(* IEC 61131-3 sources: plcassist-cli/packages/volt-lsp-iec/test-corpus/bakon-nano/Device/Plc Logic/Application/Library Manager/L_TP2P_TechModulesProcessFunctions, 25 files *)

(* ---- GETBOOLEANPROPERTY.fun ---- *)
FUNCTION GETBOOLEANPROPERTY : BOOL
VAR_INPUT
	STKEY : WSTRING;
END_VAR
END_FUNCTION

(* ---- GETCOMPANY.fun ---- *)
FUNCTION GETCOMPANY : WSTRING
END_FUNCTION

(* ---- GETNUMBERPROPERTY.fun ---- *)
FUNCTION GETNUMBERPROPERTY : DINT
VAR_INPUT
	STKEY : WSTRING;
END_VAR
END_FUNCTION

(* ---- GETTEXTPROPERTY.fun ---- *)
FUNCTION GETTEXTPROPERTY : WSTRING
VAR_INPUT
	STKEY : WSTRING;
END_VAR
END_FUNCTION

(* ---- GETTEXTPROPERTY2.fun ---- *)
FUNCTION GETTEXTPROPERTY2 : POINTER TO WSTRING
VAR_INPUT
	STKEY : WSTRING;
END_VAR
END_FUNCTION

(* ---- GETTITLE.fun ---- *)
FUNCTION GETTITLE : WSTRING
END_FUNCTION

(* ---- GETVERSION.fun ---- *)
FUNCTION GETVERSION : VERSION
END_FUNCTION

(* ---- GETVERSIONPROPERTY.fun ---- *)
FUNCTION GETVERSIONPROPERTY : VERSION
VAR_INPUT
	STKEY : WSTRING;
END_VAR
END_FUNCTION

(* ---- L_TP2P_TC_CELSIUSTOFAHRENHEIT_ABS.fun ---- *)
FUNCTION L_TP2P_TC_CELSIUSTOFAHRENHEIT_ABS : LREAL
VAR_INPUT
	LRINVAL : LREAL;
END_VAR
END_FUNCTION

(* ---- L_TP2P_TC_CELSIUSTOFAHRENHEIT_REL.fun ---- *)
FUNCTION L_TP2P_TC_CELSIUSTOFAHRENHEIT_REL : LREAL
VAR_INPUT
	LRINVAL : LREAL;
END_VAR
END_FUNCTION

(* ---- _TM_COMMONBASE.fb ---- *)
FUNCTION_BLOCK _TM_COMMONBASE EXTENDS L_TB2P_TM_Base
VAR
	XTMSTOP : BOOL;
	LWTCHECKSUM : LWORD;
	ERRORHANDLER : L_IE1P_ErrorHandler;
	PINPUTBASE : POINTER TO L_TP2P_TemperatureControlBaseIn;
	POUTPUTBASE : POINTER TO L_TP2P_TemperatureControlBaseOut;
END_VAR
END_FUNCTION_BLOCK

METHOD CALL_ALLOCPOINTADR
END_METHOD

METHOD CALL_CHECKREQUESTS
END_METHOD

METHOD CALL_CTRLREQACTIVE : BOOL
END_METHOD

METHOD CALL_OUTPUT
END_METHOD

METHOD CALL_REQUESTS_EXT
END_METHOD

METHOD CALL_RESETCOMMANDS
END_METHOD

METHOD CALL_RESETOUTPUT
END_METHOD

METHOD CALL_RESETSETERROR
END_METHOD

METHOD CALL_SETERROR
END_METHOD

METHOD CALL_STOP
END_METHOD

METHOD CALL_TMFUNCTIONALITY
END_METHOD

METHOD CALL_S000_CYCLIC
END_METHOD

METHOD CALL_S001_INIT
END_METHOD

METHOD CALL_S002_READY
END_METHOD

METHOD CALL_S996_STOP
END_METHOD

METHOD CALL_STATEMACHINE
END_METHOD

METHOD CALL_T000_ALLSTATES
END_METHOD

METHOD CALL_T002_READY
END_METHOD

METHOD CALL_S000_CYCLIC_OUT
END_METHOD

METHOD CALL_S999_ERROR_OUT
END_METHOD

METHOD CALL_STATEMACHINE_OUT
END_METHOD

METHOD CALL_T000_ALLSTATES_OUT
END_METHOD

(* ---- _TM_TEMPERATURECONTROLBASE.fb ---- *)
FUNCTION_BLOCK _TM_TEMPERATURECONTROLBASE EXTENDS _TM_CommonBase
VAR_OUTPUT
	PPAR : POINTER TO _scPar_TM_TemperatureControlBase;
	PSF : POINTER TO _scSF_TM_TemperatureControlBase;
	PAP : POINTER TO _scAP_TM_TemperatureControlBase;
END_VAR
VAR_IN_OUT
	SCPERSISTENTDATA : L_TP2P_scPD_TemperatureControlBase;
END_VAR
VAR
	TM_TEMPERATURECONTROLCONFIG : L_TB2P_ModuleHandlerConfig;
	PINPUT : POINTER TO L_TP2P_TemperatureControlBaseIn;
	POUTPUT : POINTER TO L_TP2P_TemperatureControlBaseOut;
	_PSCPARVISU : POINTER TO _scPar_TM_TemperatureControlBase;
	SCPD_ACT : REFERENCE TO L_TP2P_scPD_TemperatureControlBase;
	LRTASKCYCLE : LREAL := 0.01;
	XNOREGULATIONPARAM : BOOL := FALSE;
	FB_TASKINFO : L_TP2P_TC_GetTaskInfo;
	FB_TEMPSETFILTER : L_TP2P_TC_TempSetFilter;
	FB_TEMPACTPROCESSING : L_TP2P_TC_TempActProcessing;
	FB_MONITORING : L_TP2P_TC_Monitoring;
	FB_PIDCONTROLLER : L_TP2P_TC_PIDController;
	FB_PARAMETERSWITCHING : L_TP2P_TC_ParameterSwitching;
	FB_PWM : L_TP2P_TC_PWM;
	FB_DIFFCTRL : L_TP2P_TC_DiffCtrl;
	FB_PARAMETERIDENTIFICATION : L_TP2P_TC_ParameterIdentification;
	SCIDENTDIAG : _sc_TM_TC_IdentDiagInfo;
END_VAR
END_FUNCTION_BLOCK

METHOD CALL_ALLOCPOINTADR
END_METHOD

METHOD CALL_CTRLREQACTIVE : BOOL
END_METHOD

METHOD CALL_ERRORHANDLER
END_METHOD

METHOD CALL_INITDONE
END_METHOD

METHOD CALL_INITROUTINE
END_METHOD

METHOD CALL_INTERNALCTRL
END_METHOD

METHOD CALL_OUTPUT
END_METHOD

METHOD CALL_OUTPUT_SF
END_METHOD

METHOD CALL_REQUESTS_EXT
END_METHOD

METHOD CALL_RESETCOMMANDS
END_METHOD

METHOD CALL_RESETOUTPUT
END_METHOD

METHOD CALL_FBMETHODS
END_METHOD

METHOD CALL_FB_DIFFCTRL
END_METHOD

METHOD CALL_FB_DIFFCTRLINPUTS
END_METHOD

METHOD CALL_FB_MONITORING
END_METHOD

METHOD CALL_FB_MONITORINGINPUTS
END_METHOD

METHOD CALL_FB_PIDCONTROLLER
END_METHOD

METHOD CALL_FB_PIDCONTROLLERINPUTS
END_METHOD

METHOD CALL_FB_PWM
END_METHOD

METHOD CALL_FB_PWMINPUTS
END_METHOD

METHOD CALL_FB_PARAMETERIDENTIFICATION
END_METHOD

METHOD CALL_FB_PARAMETERIDENTIFICATIONINPUTS
END_METHOD

METHOD CALL_FB_PARAMETERSWITCHING
END_METHOD

METHOD CALL_FB_PARAMETERSWITCHINGINPUTS
END_METHOD

METHOD CALL_FB_TEMPACTPROCESSING
END_METHOD

METHOD CALL_FB_TEMPACTPROCESSINGINPUTS
END_METHOD

METHOD CALL_FB_TEMPSETFILTER
END_METHOD

METHOD CALL_FB_TEMPSETFILTERINPUTS
END_METHOD

METHOD CALL_S000_CYCLIC
END_METHOD

METHOD CALL_S002_READY
END_METHOD

METHOD CALL_S210_CONTROL
END_METHOD

METHOD CALL_S211_REGULATION
END_METHOD

METHOD CALL_S212_IDENTIFICATION
END_METHOD

METHOD CALL_S996_STOP
END_METHOD

METHOD CALL_STATEMACHINE
END_METHOD

METHOD CALL_T002_READY
END_METHOD

(* ---- GLOBALTEXTLIST.fb ---- *)
FUNCTION_BLOCK GLOBALTEXTLIST
VAR
	M_TEXTLISTFILE : STRING(255);
	_STNAMESPACE : STRING;
END_VAR
END_FUNCTION_BLOCK

(* ---- L_TP2P_TC_DIFFCTRL.fb ---- *)
FUNCTION_BLOCK L_TP2P_TC_DIFFCTRL
VAR_INPUT
	LRTASKCYCLE : LREAL := 0.001;
	XENABLE : BOOL;
	LRCONTROLVALUE : LREAL;
END_VAR
VAR_OUTPUT
	XDIFFPOSITIVEOUT : BOOL;
	XDIFFNEGATIVEOUT : BOOL;
END_VAR
VAR_IN_OUT
	SCPAR : _scPar_TM_TemperatureControlBase;
END_VAR
VAR
	LRSIMUCONTROL_PCT : LREAL := 0.0;
	LRCTRLDIFF_PCT : LREAL;
	LRTIME_100PCT : LREAL := 0;
	LRTIME_0PCT : LREAL := 0;
	LRMINIMALONTIME_S : LREAL := 1;
	LRMINIMALOFFTIME_S : LREAL := 1;
	LRACTUALONTIME_POSITIVE_S : LREAL := 0;
	LRACTUALOFFTIME_POSITIVE_S : LREAL := 0;
	LRACTUALONTIME_NEGATIVE_S : LREAL := 0;
	LRACTUALOFFTIME_NEGATIVE_S : LREAL := 0;
	XPOSOUTLAST : BOOL := FALSE;
	XNEGOUTLAST : BOOL := FALSE;
END_VAR
END_FUNCTION_BLOCK

(* ---- L_TP2P_TC_GETTASKINFO.fb ---- *)
FUNCTION_BLOCK L_TP2P_TC_GETTASKINFO
VAR_OUTPUT
	DWCYCLETIME : DWORD;
	LRCYCLETIME : LREAL;
END_VAR
VAR
	XFIRSTCYCLE : BOOL := TRUE;
	HANDLE : RTS_IEC_HANDLE;
	INTERVAL : UDINT;
END_VAR
END_FUNCTION_BLOCK

(* ---- L_TP2P_TC_MONITORING.fb ---- *)
FUNCTION_BLOCK L_TP2P_TC_MONITORING
VAR_INPUT
	LRTASKCYCLE : LREAL := 0.001;
	XENABLE : BOOL := FALSE;
	LRSETTEMP : LREAL := 0;
	LRACTTEMP : LREAL := 0;
	LRACTTEMPUNFILTERED : LREAL := 0;
END_VAR
VAR_OUTPUT
	XTEMPMAXCRITICALABSOLUTE : BOOL;
	XSETTEMPREACHED : BOOL;
	XTEMPMIN : BOOL;
	XTEMPMAX : BOOL;
	XSENSORMONITORINGVALUEMIN : BOOL;
	XSENSORMONITORINGVALUEMAX : BOOL;
	XSENSORMONITORINGCHANGEMAX : BOOL;
END_VAR
VAR_IN_OUT
	SCPAR : _scPar_TM_TemperatureControlBase;
END_VAR
VAR
	LRSETACTDIFF : LREAL;
	LRACTTEMPLASTCYCLE : LREAL;
	RTENABLE : R_TRIG;
END_VAR
END_FUNCTION_BLOCK

(* ---- L_TP2P_TC_PARAMETERIDENTIFICATION.fb ---- *)
FUNCTION_BLOCK L_TP2P_TC_PARAMETERIDENTIFICATION
VAR_INPUT
	XENABLE : BOOL := FALSE;
	LRTASKCYCLE : LREAL := 0.001;
	LRTEMPACT : LREAL;
END_VAR
VAR_OUTPUT
	XDONE : BOOL;
	XBUSY : BOOL;
	WERRORID : WORD;
	WSTEP : WORD;
	WPHASE : WORD;
	LRCONTROLVALUEOUT : LREAL;
	LRTAUDEAD : LREAL;
	LRKI : LREAL;
	LRIDENTS1ELAPSEDTIME : LREAL;
	LRIDENTS1TEMPACTGRADIENT : LREAL;
	LRIDENTS2TEMPSTART : LREAL;
	LRIDENTS2ELAPSEDTIME : LREAL;
	LRIDENTS2TEMPACTGRADIENT : LREAL;
	LRIDENTS3TAUDEADACT : LREAL;
	LRIDENTS3TAUDEADMAX : LREAL;
END_VAR
VAR_IN_OUT
	SCPAR : _scPar_TM_TemperatureControlBase;
	SCPD : L_TP2P_scPD_TemperatureControlBase;
	SCIDENTDIAG : _sc_TM_TC_IdentDiagInfo;
END_VAR
VAR
	DWREGDATASIZE : DWORD := 20;
	FB_TEMPACTT1 : L_TP2P_TC_PT1Process;
	LRTEMPACTVALUE : LREAL;
	LRTEMPACTGRADIENT : LREAL;
	LRTEMPACTLASTCYCLE : LREAL;
	LRTIMESTART_S1 : LREAL;
	LRTEMPSTART_S2 : LREAL;
	LRTIMESTART_S2 : LREAL;
	LRTEMPSTART_S3 : LREAL;
	LRTIMESTART_S3 : LREAL;
	LRCONTROLVALUESTART_S3 : LREAL;
	LRCONTROLVALUESTEP_S3 : LREAL;
	DICYCLECOUNT_S3 : DINT;
	UDIREG_N : UDINT;
	LRREG_SUMX : LREAL;
	LRREG_SUMY : LREAL;
	LRREG_SUMXX : LREAL;
	LRREG_SUMXY : LREAL;
	LRREG_XM : LREAL;
	LRREG_YM : LREAL;
	LRREG_A : LREAL;
	LRREG_B : LREAL;
	LRZAEHLER_B : LREAL;
	LRNENNER_B : LREAL;
	LRTAUDEADMAX : LREAL;
	LRTAUDEADACT : LREAL;
	LRBMAX : LREAL;
	LRPAR_STEP1TEMPCHANGEMAX : LREAL;
	LRPAR_STEP2CONTROLSTEPPCT : LREAL;
	LRPAR_STEP2TEMPCHANGEMAX : LREAL;
	LRPAR_STEP2TEMPDIFFMIN : LREAL;
	LRPAR_STEP2WAITTIMEMIN : LREAL;
	LRPAR_STEP2CONTROLVALUEMAXPCT : LREAL;
	LRPAR_STEP3CONTROLSTEPPCT : LREAL;
	LRPAR_STEP3TEMPDIFFMIN : LREAL;
	LRPAR_STEP3REGRESSIONTIME : LREAL;
	ALRXVAL : ARRAY [1..dwRegDataSize] OF LREAL;
	ALRYVAL : ARRAY [1..dwRegDataSize] OF LREAL;
	DWCNT : DWORD;
	XPERFORMCALCREGRESSION : BOOL := FALSE;
	LRR01 : LREAL;
	LRSAMPLETIME : LREAL := 0.1;
	LRBUFFERLENGTH : LREAL := 0;
END_VAR
END_FUNCTION_BLOCK

METHOD ADDREGPOINT
VAR_INPUT
	LRX : LREAL;
	LRY : LREAL;
END_VAR
END_METHOD

METHOD CALCREGRESSION
END_METHOD

METHOD PREPAREREGBUFFER
END_METHOD

METHOD RESET : BOOL
END_METHOD

(* ---- L_TP2P_TC_PARAMETERIDENTIFICATION_T30.fb ---- *)
FUNCTION_BLOCK L_TP2P_TC_PARAMETERIDENTIFICATION_T30
VAR_INPUT
	XENABLE : BOOL := FALSE;
	LRTASKCYCLE : LREAL := 0.001;
	LRTEMPACT : LREAL;
END_VAR
VAR_OUTPUT
	XDONE : BOOL;
	XBUSY : BOOL;
	WERRORID : WORD;
	WSTEP : WORD;
	WPHASE : WORD;
	LRCONTROLVALUEOUT : LREAL;
	LRTAUDEAD : LREAL;
	LRKI : LREAL;
END_VAR
VAR_IN_OUT
	SCPAR : _scPar_TM_TemperatureControlBase;
	SCPD : L_TP2P_scPD_TemperatureControlBase;
END_VAR
VAR
	DWREGDATASIZE : DWORD := 30;
	FB_TEMPACTT1 : L_TP2P_TC_PT1Process;
	LRTEMPACTVALUE : LREAL;
	LRTEMPACTGRADIENT : LREAL;
	LRTEMPACTLASTCYCLE : LREAL;
	LRTIMESTART_S1 : LREAL;
	LRTEMPSTART_S2 : LREAL;
	LRTIMESTART_S2 : LREAL;
	LRTEMPSTART_S3 : LREAL;
	LRTIMESTART_S3 : LREAL;
	LRCONTROLVALUESTART_S3 : LREAL;
	LRCONTROLVALUESTEP_S3 : LREAL;
	DICYCLECOUNT_S3 : DINT;
	UDIREG_N : UDINT;
	LRREG_SUMX : LREAL;
	LRREG_SUMY : LREAL;
	LRREG_SUMXX : LREAL;
	LRREG_SUMXY : LREAL;
	LRREG_XM : LREAL;
	LRREG_YM : LREAL;
	LRREG_A : LREAL;
	LRREG_B : LREAL;
	LRZAEHLER_B : LREAL;
	LRNENNER_B : LREAL;
	LRTAUDEADMAX : LREAL;
	LRTAUDEADACT : LREAL;
	LRBMAX : LREAL;
	LRPAR_STEP1TEMPCHANGEMAX : LREAL;
	LRPAR_STEP2CONTROLSTEPPCT : LREAL;
	LRPAR_STEP2TEMPCHANGEMAX : LREAL;
	LRPAR_STEP2TEMPDIFFMIN : LREAL;
	LRPAR_STEP2WAITTIMEMIN : LREAL;
	LRPAR_STEP2CONTROLVALUEMAXPCT : LREAL;
	LRPAR_STEP3CONTROLSTEPPCT : LREAL;
	LRPAR_STEP3TEMPDIFFMIN : LREAL;
	ALRXVAL : ARRAY [1..dwRegDataSize] OF LREAL;
	ALRYVAL : ARRAY [1..dwRegDataSize] OF LREAL;
	DWCNT : DWORD;
	XPERFORMCALCREGRESSION : BOOL := FALSE;
	LRR01 : LREAL;
END_VAR
END_FUNCTION_BLOCK

METHOD ADDREGPOINT
VAR_INPUT
	LRX : LREAL;
	LRY : LREAL;
END_VAR
END_METHOD

METHOD CALCREGRESSION
END_METHOD

METHOD PREPAREREGBUFFER
END_METHOD

(* ---- L_TP2P_TC_PARAMETERSWITCHING.fb ---- *)
FUNCTION_BLOCK L_TP2P_TC_PARAMETERSWITCHING
VAR_INPUT
	XENABLE : BOOL := FALSE;
	LRTASKCYCLE : LREAL := 0.001;
	LRSETVALUE : LREAL;
	LRACTVALUE : LREAL;
	LRDEVIATIONCONSTRAINTA : LREAL;
	LRDEVIATIONCONSTRAINTB : LREAL;
	LRGAINFACTORDISTURBANCECONTROL : LREAL;
	LRFILTERTIMEFACTORDISTURBANCECONTROL : LREAL;
	LRGAINFACTORREFERENCECONTROL : LREAL;
	LRFILTERTIMEFACTORREFERENCECONTROL : LREAL;
	LRGAINORIGINAL : LREAL;
	LRTEMPSETFILTERTIMEORIGINAL : LREAL;
END_VAR
VAR_OUTPUT
	XREFERENCECONTROLACTIVE : BOOL;
	XDISTURBANCECONTROLACTIVE : BOOL;
	LRGAINACTUAL : LREAL;
	LRTEMPSETFILTERTIMEACTUAL : LREAL;
END_VAR
VAR_IN_OUT
	SCPAR : _scPar_TM_TemperatureControlBase;
END_VAR
END_FUNCTION_BLOCK

(* ---- L_TP2P_TC_PIDCONTROLLER.fb ---- *)
FUNCTION_BLOCK L_TP2P_TC_PIDCONTROLLER
VAR_INPUT
	XENABLE : BOOL := FALSE;
	LRTASKCYCLE : LREAL := 0.001;
	LRSETVALUE : LREAL;
	LRACTVALUE : LREAL;
	LRGAIN : LREAL;
	LRINTEGRALTIME : LREAL;
	LRDERIVATIVETIME : LREAL;
END_VAR
VAR_OUTPUT
	LRCONTROLVALUE : LREAL;
	XCONTROLVALUELIMITATIONACTIVE : BOOL;
	LRPVALUE : LREAL;
	LRIVALUE : LREAL;
	LRDVALUE : LREAL;
	LRCONTROLVALUEUNLIMITED : LREAL;
END_VAR
VAR_IN_OUT
	SCPAR : _scPar_TM_TemperatureControlBase;
END_VAR
VAR
	LRTEMPDIFF : LREAL := 0;
	LRINTEGRALSUM : LREAL := 0;
	XICLAMPINGACTIVE : BOOL;
	DPT1 : L_TP2P_TC_PT1Process;
	LRTEMPDIFFFILTERED : LREAL;
	XFIRSTENABLEDCYCLE : BOOL := TRUE;
	LRTEMPDIFFLASTCYCLE : LREAL;
	LRRP1 : LREAL;
	XXP1 : BOOL;
END_VAR
END_FUNCTION_BLOCK

(* ---- L_TP2P_TC_PT1PROCESS.fb ---- *)
FUNCTION_BLOCK L_TP2P_TC_PT1PROCESS
VAR_INPUT
	LRKP : LREAL := 200;
	LRT1 : LREAL := 2;
	LRTASKCYCLE : LREAL := 0.001;
	XT1ZERO : BOOL := FALSE;
	LRINVAL : LREAL := 0;
END_VAR
VAR_OUTPUT
	LROUTVAL : LREAL := 0;
END_VAR
VAR
	LROUTTARGET : LREAL := 0;
END_VAR
END_FUNCTION_BLOCK

(* ---- L_TP2P_TC_PWM.fb ---- *)
FUNCTION_BLOCK L_TP2P_TC_PWM
VAR_INPUT
	LRTASKCYCLE : LREAL := 0.001;
	XENABLE : BOOL;
	LRCONTROLVALUE : LREAL;
END_VAR
VAR_OUTPUT
	LRHEATINGPOWERPCT : LREAL;
	LRHEATINGPOWERSCALED : LREAL;
	XPWMOUT : BOOL;
END_VAR
VAR_IN_OUT
	SCPAR : _scPar_TM_TemperatureControlBase;
END_VAR
VAR
	LRCVNOM : LREAL := 0.0;
	LRCVACT : LREAL;
	DNCVACTTICKS : DINT;
	DNCVPWMTICKS : DINT;
	LRCVREST : LREAL := 0;
	LRCVRESOLUTION : LREAL;
END_VAR
END_FUNCTION_BLOCK

(* ---- L_TP2P_TC_TEMPACTPROCESSING.fb ---- *)
FUNCTION_BLOCK L_TP2P_TC_TEMPACTPROCESSING
VAR_INPUT
	LRTASKCYCLE : LREAL := 0.001;
	LRACTSENSORIN : LREAL := 0;
	LRPT1TIMEDELAY : LREAL := 30;
END_VAR
VAR_OUTPUT
	LRTEMPACTUNFILTERED : LREAL := 0;
	LRTEMPACT : LREAL := 0;
END_VAR
VAR_IN_OUT
	SCPAR : _scPar_TM_TemperatureControlBase;
END_VAR
VAR
	FB_PT1 : L_TP2P_TC_PT1Process;
	LRSENSORVALWITHGAIN : LREAL;
	LRSENSORVALWITHOFFSET : LREAL;
END_VAR
END_FUNCTION_BLOCK

(* ---- L_TP2P_TC_TEMPSETFILTER.fb ---- *)
FUNCTION_BLOCK L_TP2P_TC_TEMPSETFILTER
VAR_INPUT
	LRTASKCYCLE : LREAL := 0.001;
	XENABLE : BOOL := FALSE;
	LRPT1TIMEDELAY : LREAL := 30;
	LRSETPOINTIN : LREAL := 0;
	LROUTVALUEIFDISABLED : LREAL := 0;
END_VAR
VAR_OUTPUT
	XENABLED : BOOL := FALSE;
	LRSETPOINTOUT : LREAL := 0;
	XFILTERACTIVE : BOOL := FALSE;
END_VAR
VAR_IN_OUT
	SCPAR : _scPar_TM_TemperatureControlBase;
END_VAR
VAR
	LRSETPOINTINLAST : LREAL := 0;
	RTENABLE : R_TRIG;
	FBPT1 : L_TP2P_TC_PT1Process;
	LRCALC01 : LREAL;
END_VAR
END_FUNCTION_BLOCK

(* ---- L_TP2P_TEMPERATURECONTROLBASE.fb ---- *)
FUNCTION_BLOCK L_TP2P_TEMPERATURECONTROLBASE EXTENDS L_TB2P_TechModuleBase
VAR_INPUT
	XENABLEINTERNALCONTROL : BOOL;
	XENABLE : BOOL;
	XRESETERROR : BOOL;
	XSTOP : BOOL;
	XTEMPERATURECTRL : BOOL;
	XIDENTCTRLPAR : BOOL;
	LRSETTEMP : LREAL;
	SCPAR : L_TP2P_scPar_TemperatureControlBase;
	SCACCESSPOINTS : L_TP2P_scAP_TemperatureControlBase;
	NACTSENSORIN : INT;
END_VAR
VAR_OUTPUT
	ETMSTATE : L_TP2P_States := L_TP2P_States.INIT;
	XERROR : BOOL;
	XWARNING : BOOL;
	EERRORID : L_IE1P_Error;
	SCSIGNALFLOW : L_TP2P_scSF_TemperatureControlBase;
	LRACTTEMP : LREAL;
	XPWMOUT : BOOL;
	XDIFFPOSITIVEOUT : BOOL;
	XDIFFNEGATIVEOUT : BOOL;
	LRHEATINGPOWERPCT : LREAL;
	LRHEATINGPOWERSCALED : LREAL;
	WIDENTPHASE : WORD;
	XIDENTBUSY : BOOL;
	XIDENTDONE : BOOL;
	XTEMPMAX : BOOL;
	XTEMPMIN : BOOL;
	XSETTEMPREACHED : BOOL;
END_VAR
VAR_IN_OUT
	SCPERSISTENTDATA : L_TP2P_scPD_TemperatureControlBase;
END_VAR
VAR
	TM_INT : _TM_TemperatureControlBase := STRUCT(ModuleHandler := ModuleHandler);
	SCPAR_INT : L_TP2P_scPar_TemperatureControlBase;
	XENABLEOLD : BOOL;
	_UICALLMFUNIDXINPUT : UINT := 1;
	_UICALLMFUNIDXOUTPUT : UINT := 1;
	_ASCINPUT : ARRAY [1.._MCCall.c_BufferDepthInput] OF L_TP2P_TemperatureControlBaseIn;
	_ASCOUTPUT : ARRAY [1.._MCCall.c_BufferDepthOutput] OF L_TP2P_TemperatureControlBaseOut;
	_ASCPARCORE : ARRAY [1.._MCCall.c_BufferDepthInput] OF L_TP2P_scPar_TemperatureControlBase;
	_MCCALL : L_UM1P_MCCall;
	_ASCACCESSPOINTSCORE : ARRAY [1.._MCCall.c_BufferDepthInput] OF L_TP2P_scAP_TemperatureControlBase;
	_ASCSIGNALFLOWCORE : ARRAY [1.._MCCall.c_BufferDepthOutput] OF L_TP2P_scSF_TemperatureControlBase;
	_SCINPUTVISU : L_TP2P_TemperatureControlBaseIn;
	_PSCINPUTVISU : POINTER TO L_TP2P_TemperatureControlBaseIn := ADR(_scInputVisu);
	_PSCOUTPUTVISU : POINTER TO L_TP2P_TemperatureControlBaseOut := ADR(_ascOutput[1]);
	_PSCPARVISU : POINTER TO L_TP2P_scPar_TemperatureControlBase := ADR(scPar_int);
	ITFITECHMODULEINTERNAL : L_TB2P_ITechModuleInternal;
END_VAR
END_FUNCTION_BLOCK

METHOD GET_PAP : POINTER TO L_TB2P_scAP_TM_MotionControl
END_METHOD

METHOD GET_PPAR : POINTER TO L_TB2P_scPar_TM_MotionControl
END_METHOD

METHOD GET_PSF : POINTER TO L_TB2P_scSF_TM_MotionControl
END_METHOD

METHOD CALLFUNCTION
VAR_INPUT
	UIINPUTDATAIDX : UINT;
	UIOUTPUTDATAIDX : UINT;
END_VAR
END_METHOD

METHOD COPYINPUTS : BOOL
VAR_INPUT
	IDX : WORD;
END_VAR
END_METHOD

METHOD COPYOUTPUTS : BOOL
VAR_INPUT
	IDX : WORD;
END_VAR
END_METHOD

METHOD FUNCTIONWASCALLEDTWICE : BOOL
VAR_INPUT
	IDX : WORD;
END_VAR
END_METHOD

METHOD HANDLESTANDARDCALL : BOOL
END_METHOD

METHOD SYNCOUTPUTS
VAR_INPUT
	UICOPYOUTPUTFROMIDX : UINT;
	UICOPYOUTPUTTOIDX : UINT;
END_VAR
END_METHOD

METHOD CALL_INTERNALCTRL
END_METHOD
